Fanuc KAREL source: KX00026.KL

PROGRAM KX00026
%NOLOCKGROUP
%PRIORITY = 20
VAR
  I: INTEGER
  J: INTEGER
  B: BOOLEAN
  F: FILE
  S: STRING[80]
  P: XYZWPR
BEGIN
  I = 1
END KX00026
